(* IEC 61131-3 sources: llm-plc-st-eval/data/definitivo/gemini-3.1-pro-preview/B4/few_shot, 3 files *)

(* ---- ejec_1.st ---- *)
FUNCTION_BLOCK FB_Giro
VAR_INPUT
    btnFwd : BOOL; (* Boton de giro horario *)
    btnRev : BOOL; (* Boton de giro antihorario *)
    btnParo : BOOL; (* Boton de paro *)
END_VAR
VAR_OUTPUT
    fwd : BOOL; (* Salida de giro horario *)
    rev : BOOL; (* Salida de giro antihorario *)
END_VAR

(* Enclavamiento de giro horario: requiere que no este activo el paro ni el giro inverso *)
fwd := (btnFwd OR fwd) AND NOT btnParo AND NOT rev;

(* Enclavamiento de giro antihorario: requiere que no este activo el paro ni el giro horario *)
rev := (btnRev OR rev) AND NOT btnParo AND NOT fwd;
END_FUNCTION_BLOCK

(* ---- ejec_2.st ---- *)
FUNCTION_BLOCK FB_Giro
VAR_INPUT
    btnFwd : BOOL; (* Boton de marcha en sentido horario *)
    btnRev : BOOL; (* Boton de marcha en sentido antihorario *)
    btnParo : BOOL; (* Boton de paro *)
END_VAR
VAR_OUTPUT
    fwd : BOOL; (* Salida para giro horario *)
    rev : BOOL; (* Salida para giro antihorario *)
END_VAR

(* Enclavamiento para giro horario: requiere que no este activo el paro ni el giro opuesto *)
fwd := (fwd OR btnFwd) AND NOT btnParo AND NOT rev;

(* Enclavamiento para giro antihorario: requiere que no este activo el paro ni el giro opuesto *)
rev := (rev OR btnRev) AND NOT btnParo AND NOT fwd;
END_FUNCTION_BLOCK

(* ---- ejec_3.st ---- *)
FUNCTION_BLOCK FB_Giro
VAR_INPUT
    btnFwd : BOOL; (* Boton de giro horario *)
    btnRev : BOOL; (* Boton de giro antihorario *)
    btnParo : BOOL; (* Boton de paro *)
END_VAR
VAR_OUTPUT
    fwd : BOOL; (* Salida de giro horario *)
    rev : BOOL; (* Salida de giro antihorario *)
END_VAR

(* Enclavamiento de giro horario: requiere que no este activo el paro ni el giro opuesto *)
fwd := (btnFwd OR fwd) AND NOT btnParo AND NOT rev;

(* Enclavamiento de giro antihorario: requiere que no este activo el paro ni el giro opuesto *)
rev := (btnRev OR rev) AND NOT btnParo AND NOT fwd;
END_FUNCTION_BLOCK
